(* IEC 61131-3 sources: Lasal-MCP/examples/SampleSource/4_PumpControlSchemeSolution/Stations/MachineControl/MachineControl/Class/_EventAddfromPLC, 1 file *)

(* ---- _EventAddfromPLC.st ---- *)
#ifndef EVENT_VALUECHANGE
  #define   Event_ValueChange               16#102      // Event für: Variable vom Typ Numeric
#endif

#ifndef EVENT_EVENTENTRY
  #define   Event_EventEntry                16#270
#endif

(*!
<Class
	Name               = "_EventAddfromPLC"
	Revision           = "1.4"
	RealtimeTask       = "false"
	CyclicTask         = "true"
	BackgroundTask     = "true"
	Sigmatek           = "true"
	OSInterface        = "false"
	HighPriority       = "false"
	Automatic          = "false"
	UpdateMode         = "Prescan"
	SharedCommandTable = "true"
	Objectsize         = "(470,120)"
	Comment            = "class for adding an event from plc and sending it to HMI via DataManager">
	<Channels>
		<Server Name="ClassSvr">
			<NewInst>
				<Function Name="NewInst_AddSystemOnOff">
					<InputParameter>
						<Parameter Name="dDate"/>
						<Parameter Name="dTime"/>
						<Parameter Name="bSwitchOnOff"/>
					</InputParameter>
					<OutputParameter>
						<Parameter Name="ret_code"/>
					</OutputParameter>
				</Function>
				<Function Name="NewInst_AddEventEntry">
					<InputParameter>
						<Parameter Name="config"/>
						<Parameter Name="uiCategory"/>
						<Parameter Name="uiIndex"/>
						<Parameter Name="pText"/>
						<Parameter Name="uiSize"/>
						<Parameter Name="bUnicode"/>
					</InputParameter>
					<OutputParameter>
						<Parameter Name="ret_code"/>
					</OutputParameter>
				</Function>
				<Function Name="NewInst_AddDateChange">
					<InputParameter>
						<Parameter Name="udVarNo"/>
						<Parameter Name="dOldDate"/>
						<Parameter Name="dNewDate"/>
					</InputParameter>
					<OutputParameter>
						<Parameter Name="ret_code"/>
					</OutputParameter>
				</Function>
				<Function Name="NewInst_AddTimeChange">
					<InputParameter>
						<Parameter Name="udVarNo"/>
						<Parameter Name="dOldTime"/>
						<Parameter Name="dNewTime"/>
					</InputParameter>
					<OutputParameter>
						<Parameter Name="ret_code"/>
					</OutputParameter>
				</Function>
				<Function Name="NewInst_AddMenuChange">
					<InputParameter>
						<Parameter Name="udVarNo"/>
						<Parameter Name="udMenuIndex"/>
						<Parameter Name="dOldValue"/>
						<Parameter Name="dNewValue"/>
					</InputParameter>
					<OutputParameter>
						<Parameter Name="ret_code"/>
					</OutputParameter>
				</Function>
				<Function Name="NewInst_AddValueChange">
					<InputParameter>
						<Parameter Name="udLasalID"/>
						<Parameter Name="dOldValue"/>
						<Parameter Name="dNewValue"/>
					</InputParameter>
					<OutputParameter>
						<Parameter Name="ret_code"/>
					</OutputParameter>
				</Function>
				<Function Name="NewInst_AddOPChange">
					<InputParameter>
						<Parameter Name="eOPMode"/>
					</InputParameter>
					<OutputParameter>
						<Parameter Name="ret_code"/>
					</OutputParameter>
				</Function>
				<Function Name="NewInst_AddUserLoginLogout">
					<InputParameter>
						<Parameter Name="pUserName"/>
						<Parameter Name="dActLevel"/>
						<Parameter Name="bIsLogin"/>
					</InputParameter>
					<OutputParameter>
						<Parameter Name="ret_code"/>
					</OutputParameter>
				</Function>
			</NewInst>
		</Server>
	</Channels>
	<Dependencies>
		<Files>
			<File Path=".\Class\_EventAddfromPLC\_EventAddfromPLC_de.pdf"/>
			<File Path=".\Class\_EventAddfromPLC\_EventAddfromPLC_en.pdf"/>
		</Files>
	</Dependencies>
	<RevDoku>
		<Owner Company="Sigmatek"/>
		<Dokumentation Revision="1.4" Date="2016-10-21" Author="KaiAnd" Company="Sigmatek" Description="implemented NewInst_AddXY (Cmd 00 to Cmd 07) for adding events from external via command channel"/>
		<Dokumentation Revision="1.3" Date="2016-10-10" Author="HubChr" Company="Sigmatek" Description="Added documentation pdfs."/>
		<Dokumentation Revision="1.2" Date="2016-09-21" Author="HubChr" Company="Sigmatek" Description="Events from PLC can now also open MessageBoxes"/>
		<Dokumentation Revision="1.1" Date="2016-09-15" Author="HubChr" Company="Sigmatek" Description="Translated comments for library compatibility"/>
		<Dokumentation Revision="1.0" Date="2015-09-22" Company="Sigmatek" Description="Creation."/>
	</RevDoku>
	<Network Name="_EventAddfromPLC">
		<!-- List of Components in this network -->
		<Components>
			<Object
				Name       = "_base"
				Class      = "TCPComSend"
				Position   = "(218,120)"
				Visualized = "false">
				<Channels>
					<Server Name="ClassSvr"/>
					<Server Name="ID_Destination"/>
					<Server Name="ID_Source"/>
					<Server Name="sSendCnt"/>
					<Server Name="sSendErr"/>
					<Client Name="cPrio"/>
					<Client Name="cSendErr"/>
					<Client Name="cSendOk"/>
					<Client Name="toDataManager"/>
				</Channels>
			</Object>
		</Components>
		<Comments>
		</Comments>
		<!-- List of Connections in this network -->
		<Connections>
			<Connection Source="this.ClassSvr" Destination="_base.ClassSvr" Vertices="(1006,210),(834,210),"/>
			<Connection Source="this.ID_Destination" Destination="_base.ID_Destination" Vertices="(1006,270),(834,270),"/>
			<Connection Source="this.ID_Source" Destination="_base.ID_Source" Vertices="(1006,330),(834,330),"/>
			<Connection Source="this.sSendCnt" Destination="_base.sSendCnt" Vertices="(1006,390),(834,390),"/>
			<Connection Source="this.sSendErr" Destination="_base.sSendErr" Vertices="(1006,450),(834,450),"/>
			<Connection Source="_base.toDataManager" Destination="this.toDataManager" Vertices="(218,210),(38,210),"/>
			<Connection Source="_base.cPrio" Destination="this.cPrio" Vertices="(218,270),(38,270),"/>
		</Connections>
		<!-- Headerfiles -->
		<Options>
		</Options>
	</Network>
</Class>
*)
#pragma using TCPComSend

_EventAddfromPLC : CLASS
: TCPComSend
	TYPE
#pragma pack(push, 1)
	  _PLCEventdata : STRUCT
	    EventType : UINT;
	    no_para : UINT;
	    Para1 : DINT;
	    Para2 : DINT;
	    Para3 : DINT;
	    Para4 : DINT;
	    Para5 : DINT;
	    Para6 : DINT;
	    Para7 : DINT;
	    Para8 : DINT;
	    StringSize : UINT;
	    aString : ARRAY [0..24] OF DINT;
	  END_STRUCT;
#pragma pack(pop)
	  CmdClassSvr :  //! <Type Public="true" Name="CmdClassSvr"/>
	  (
	    NewInst_AddSystemOnOff:=0,
	    NewInst_AddEventEntry,
	    NewInst_AddDateChange,
	    NewInst_AddTimeChange,
	    NewInst_AddMenuChange,
	    NewInst_AddValueChange,
	    NewInst_AddOPChange,
	    NewInst_AddUserLoginLogout
	  )$UINT;
	END_TYPE
  //Servers:
  //Clients:
  //Variables:
  //Functions:
				//! <Function Comment="Initialization of the eventdata." Name="InitPLCEventdata"/>
	FUNCTION InitPLCEventdata
		VAR_INPUT
			pPLCEvent 	: ^_PLCEventdata;			//! <Variable Comment="Pointer to the event data." Name="InitPLCEventdata.pPLCEvent"/>
		END_VAR;
				//! <Function Comment="Sends an event for a value change to the remote station." Name="AddValueChange"/>
	FUNCTION GLOBAL AddValueChange
		VAR_INPUT
			udLasalID 	: UDINT;			//! <Variable Comment="Lasal-ID" Name="AddValueChange.udLasalID"/>
			dOldValue 	: DINT;			//! <Variable Comment="Old value" Name="AddValueChange.dOldValue"/>
			dNewValue 	: DINT;			//! <Variable Comment="New value" Name="AddValueChange.dNewValue"/>
		END_VAR;
				//! <Function Comment="Method for sending the data of a event to the remote station." Name="AddEventEntry"/>
	FUNCTION GLOBAL AddEventEntry
		VAR_INPUT
			config 	: BDINT;			//! <Variable Comment="Category for the event:&#13;&#10;0 .. System category 1&#13;&#10;1 .. System category 2&#13;&#10;2 .. System category 3&#13;&#10;3 .. System category 4&#13;&#10;4 .. Change of the OP mode&#13;&#10;else .. System category 1" Name="AddEventEntry.config"/>
			uiCategory 	: UINT;			//! <Variable Comment="Category for the event:&#13;&#10;0 .. System category 1&#13;&#10;1 .. System category 2&#13;&#10;2 .. System category 3&#13;&#10;3 .. System category 4&#13;&#10;4 .. Change of the OP mode&#13;&#10;else .. System category 1" Name="AddEventEntry.uiCategory"/>
			uiIndex 	: UINT;			//! <Variable Comment="Index in the textscheme (if used).&#13;&#10;Note: If event is for example a menue-change -&gt; menue-index." Name="AddEventEntry.uiIndex"/>
			pText 	: ^void;			//! <Variable Comment="Individual text" Name="AddEventEntry.pText"/>
			uiSize 	: UINT;			//! <Variable Comment="Size of the text" Name="AddEventEntry.uiSize"/>
			bUnicode 	: BOOL;			//! <Variable Comment="Character size of the string:&#13;&#10;FALSE .. ASCII&#13;&#10;TRUE .. UNI-Code" Name="AddEventEntry.bUnicode"/>
		END_VAR;

	FUNCTION ClassSvr::NewInst_AddSystemOnOff
		VAR_INPUT
			dDate 	: DINT;
			dTime 	: DINT;
			bSwitchOnOff 	: DINT;
		END_VAR
		VAR_OUTPUT
			ret_code 	: IprStates;
		END_VAR;

	FUNCTION ClassSvr::NewInst_AddEventEntry
		VAR_INPUT
			config 	: DINT;
			uiCategory 	: DINT;
			uiIndex 	: DINT;
			pText 	: DINT;
			uiSize 	: DINT;
			bUnicode 	: DINT;
		END_VAR
		VAR_OUTPUT
			ret_code 	: IprStates;
		END_VAR;

	FUNCTION ClassSvr::NewInst_AddDateChange
		VAR_INPUT
			udVarNo 	: DINT;
			dOldDate 	: DINT;
			dNewDate 	: DINT;
		END_VAR
		VAR_OUTPUT
			ret_code 	: IprStates;
		END_VAR;

	FUNCTION ClassSvr::NewInst_AddTimeChange
		VAR_INPUT
			udVarNo 	: DINT;
			dOldTime 	: DINT;
			dNewTime 	: DINT;
		END_VAR
		VAR_OUTPUT
			ret_code 	: IprStates;
		END_VAR;

	FUNCTION ClassSvr::NewInst_AddMenuChange
		VAR_INPUT
			udVarNo 	: DINT;
			udMenuIndex 	: DINT;
			dOldValue 	: DINT;
			dNewValue 	: DINT;
		END_VAR
		VAR_OUTPUT
			ret_code 	: IprStates;
		END_VAR;

	FUNCTION ClassSvr::NewInst_AddValueChange
		VAR_INPUT
			udLasalID 	: DINT;
			dOldValue 	: DINT;
			dNewValue 	: DINT;
		END_VAR
		VAR_OUTPUT
			ret_code 	: IprStates;
		END_VAR;

	FUNCTION ClassSvr::NewInst_AddOPChange
		VAR_INPUT
			eOPMode 	: DINT;
		END_VAR
		VAR_OUTPUT
			ret_code 	: IprStates;
		END_VAR;

	FUNCTION ClassSvr::NewInst_AddUserLoginLogout
		VAR_INPUT
			pUserName 	: DINT;
			dActLevel 	: DINT;
			bIsLogin 	: DINT;
		END_VAR
		VAR_OUTPUT
			ret_code 	: IprStates;
		END_VAR;
				//! <Function Name="ClassSvr.NewInst" Hidden="true"/>
	FUNCTION VIRTUAL GLOBAL ClassSvr::NewInst
		VAR_INPUT
			pPara 	: ^CmdStruct;
			pResult 	: ^results;
		END_VAR
		VAR_OUTPUT
			ret_code 	: iprStates;
		END_VAR;
  //Tables:
	FUNCTION @STD
		VAR_OUTPUT
			ret_code	: CONFSTATES;
		END_VAR;
	FUNCTION GLOBAL TAB @CT_;
END_CLASS;

FUNCTION VIRTUAL GLOBAL _EventAddfromPLC::ClassSvr::NewInst
	VAR_INPUT
		pPara 	: ^CmdStruct;
		pResult 	: ^Results;
	END_VAR
	VAR_OUTPUT
		ret_code 	: IprStates;
	END_VAR
	CASE pPara^.uiCmd$CmdClassSvr OF
		NewInst_AddSystemOnOff:
			ret_code := NewInst_AddSystemOnOff(pPara^.aPara[0],pPara^.aPara[1],pPara^.aPara[2]);
			pResult^.uiLng := 0 + sizeof(pResult^.uiLng);
		NewInst_AddEventEntry:
			ret_code := NewInst_AddEventEntry(pPara^.aPara[0],pPara^.aPara[1],pPara^.aPara[2],pPara^.aPara[3],pPara^.aPara[4],pPara^.aPara[5]);
			pResult^.uiLng := 0 + sizeof(pResult^.uiLng);
		NewInst_AddDateChange:
			ret_code := NewInst_AddDateChange(pPara^.aPara[0],pPara^.aPara[1],pPara^.aPara[2]);
			pResult^.uiLng := 0 + sizeof(pResult^.uiLng);
		NewInst_AddTimeChange:
			ret_code := NewInst_AddTimeChange(pPara^.aPara[0],pPara^.aPara[1],pPara^.aPara[2]);
			pResult^.uiLng := 0 + sizeof(pResult^.uiLng);
		NewInst_AddMenuChange:
			ret_code := NewInst_AddMenuChange(pPara^.aPara[0],pPara^.aPara[1],pPara^.aPara[2],pPara^.aPara[3]);
			pResult^.uiLng := 0 + sizeof(pResult^.uiLng);
		NewInst_AddValueChange:
			ret_code := NewInst_AddValueChange(pPara^.aPara[0],pPara^.aPara[1],pPara^.aPara[2]);
			pResult^.uiLng := 0 + sizeof(pResult^.uiLng);
		NewInst_AddOPChange:
			ret_code := NewInst_AddOPChange(pPara^.aPara[0]);
			pResult^.uiLng := 0 + sizeof(pResult^.uiLng);
		NewInst_AddUserLoginLogout:
			ret_code := NewInst_AddUserLoginLogout(pPara^.aPara[0],pPara^.aPara[1],pPara^.aPara[2]);
			pResult^.uiLng := 0 + sizeof(pResult^.uiLng);
	ELSE

	ret_code := READY;
	END_CASE;

END_FUNCTION

FUNCTION _EventAddfromPLC::InitPLCEventdata
	VAR_INPUT
		pPLCEvent 	: ^_PLCEventdata;
	END_VAR

  pPLCEvent^.EventType  := 0;
  pPLCEvent^.no_para    := 0;
  pPLCEvent^.Para1      := 0;
  pPLCEvent^.Para2      := 0;
  pPLCEvent^.Para3      := 0;
  pPLCEvent^.Para4      := 0;
  pPLCEvent^.Para5      := 0;
  pPLCEvent^.Para6      := 0;
  pPLCEvent^.Para7      := 0;
  pPLCEvent^.Para8      := 0;
  pPLCEvent^.StringSize := 0;
  _memset(dest := #pPLCEvent^.aString[0], usByte:=0, cntr:=sizeof(pPLCEvent^.aString));

END_FUNCTION

FUNCTION GLOBAL _EventAddfromPLC::AddValueChange
	VAR_INPUT
		udLasalID : UDINT;
		dOldValue : DINT;
		dNewValue : DINT;
	END_VAR
  VAR
  	tmpEvent : _PLCEventdata;
  END_VAR

  InitPLCEventdata(pPLCEvent:=#tmpEvent);

  // add event for change of value
  tmpEvent.EventType := EVENT_VALUECHANGE;

  // store information
  tmpEvent.no_para := 3;
  tmpEvent.para1   := udLasalID$DINT;
  tmpEvent.para2   := dOldValue;
  tmpEvent.para3   := dNewValue;

  SendData(pData:=#tmpEvent$^void, length:=sizeof(tmpEvent), timeout:=1000, OptCMD:=0);

END_FUNCTION

FUNCTION GLOBAL _EventAddfromPLC::AddEventEntry
	VAR_INPUT
		config 	   : BDINT;
		uiCategory : UINT;
		uiIndex 	 : UINT;
		pText 	   : ^void;
		uiSize 	   : UINT;
		bUnicode 	 : BOOL;
	END_VAR
  VAR
  	tmpEvent : _PLCEventdata;
  END_VAR

  InitPLCEventdata(pPLCEvent:=#tmpEvent);

  tmpEvent.EventType := EVENT_EVENTENTRY;

  // store information
  tmpEvent.no_para := 3;
  tmpEvent.para1   := to_dint(uiCategory);
  tmpEvent.para2   := to_dint(uiIndex);
  tmpEvent.para3   := bUnicode;
  tmpEvent.para4   := config$DINT;

  if ( (pText <> NIL) & (uiSize < (sizeof(tmpEvent.aString) -1)) ) then

    tmpEvent.StringSize := uiSize;
    _memcpy(ptr1:=#tmpEvent.aString[0], ptr2:=pText, cntr:=uiSize);

  end_if;

  SendData(pData:=#tmpEvent$^void, length:=sizeof(tmpEvent), timeout:=1000, OptCMD:=0);

END_FUNCTION

//***********************************************************************************************************
//  NewInst Commands for external actions via command channel
//***********************************************************************************************************

//-------------------------------------------------------------------------------------------------
//  Cmd 00: AddSystemOnOff
//-------------------------------------------------------------------------------------------------
#pragma warning(disable:73);
FUNCTION _EventAddfromPLC::NewInst_AddSystemOnOff
	VAR_INPUT
		dDate 	: DINT;
		dTime 	: DINT;
		bSwitchOnOff 	: DINT;
	END_VAR
	VAR_OUTPUT
		ret_code 	: IprStates;
	END_VAR

	ret_code := READY;

// NOT IMPLEMENTED IN PLC - reserverd for future

//  AddSystemOnOff( dDate        := dDate,
//                  dTime        := dTime,
//                  bSwitchOnOff := TO_BOOL(bSwitchOnOff) );

END_FUNCTION
#pragma warning(default:73);

//-------------------------------------------------------------------------------------------------
//  Cmd 01: AddEventEntry
//-------------------------------------------------------------------------------------------------
FUNCTION _EventAddfromPLC::NewInst_AddEventEntry
	VAR_INPUT
		config 	: DINT;
		uiCategory 	: DINT;
		uiIndex 	: DINT;
		pText 	: DINT;
		uiSize 	: DINT;
		bUnicode 	: DINT;
	END_VAR
	VAR_OUTPUT
		ret_code 	: IprStates;
	END_VAR

	ret_code := READY;

  AddEventEntry(config     := config$BDINT,
                uiCategory := TO_UINT(uiCategory),
                uiIndex    := TO_UINT(uiIndex),
                pText      := pText$^void,
                uiSize     := TO_UINT(uiSize),
                bUnicode   := TO_BOOL(bUnicode) );

END_FUNCTION

//-------------------------------------------------------------------------------------------------
//  Cmd 02: AddDateChange
//-------------------------------------------------------------------------------------------------
#pragma warning(disable:73);
FUNCTION _EventAddfromPLC::NewInst_AddDateChange
	VAR_INPUT
		udVarNo 	: DINT;
		dOldDate 	: DINT;
		dNewDate 	: DINT;
	END_VAR
	VAR_OUTPUT
		ret_code 	: IprStates;
	END_VAR

	ret_code := READY;

// NOT IMPLEMENTED IN PLC - reserverd for future

//  AddDateChange(udVarNo  := udVarNo$UDINT,
//                dOldDate := dOldDate,
//                dNewDate := dNewDate );

END_FUNCTION
#pragma warning(default:73);

//-------------------------------------------------------------------------------------------------
//  Cmd 03: AddTimeChange
//-------------------------------------------------------------------------------------------------
#pragma warning(disable:73);
FUNCTION _EventAddfromPLC::NewInst_AddTimeChange
	VAR_INPUT
		udVarNo 	: DINT;
		dOldTime 	: DINT;
		dNewTime 	: DINT;
	END_VAR
	VAR_OUTPUT
		ret_code 	: IprStates;
	END_VAR

	ret_code := READY;

// NOT IMPLEMENTED IN PLC - reserverd for future

//  AddTimeChange(udVarNo  := udVarNo$UDINT,
//                dOldTime := dOldTime,
//                dNewTime := dNewTime );

END_FUNCTION
#pragma warning(default:73);

//-------------------------------------------------------------------------------------------------
//  Cmd 04: AddMenuChange
//-------------------------------------------------------------------------------------------------
#pragma warning(disable:73);
FUNCTION _EventAddfromPLC::NewInst_AddMenuChange
	VAR_INPUT
		udVarNo 	: DINT;
		udMenuIndex 	: DINT;
		dOldValue 	: DINT;
		dNewValue 	: DINT;
	END_VAR
	VAR_OUTPUT
		ret_code 	: IprStates;
	END_VAR

	ret_code := READY;

// NOT IMPLEMENTED IN PLC - reserverd for future

//  AddMenuChange(udVarNo     := udVarNo$UDINT,
//                udMenuIndex := udMenuIndex$UDINT,
//                dOldValue   := dOldValue,
//                dNewValue   := dNewValue );

END_FUNCTION
#pragma warning(default:73);

//-------------------------------------------------------------------------------------------------
//  Cmd 05: AddValueChange
//-------------------------------------------------------------------------------------------------
FUNCTION _EventAddfromPLC::NewInst_AddValueChange
	VAR_INPUT
		udLasalID : DINT;
		dOldValue : DINT;
		dNewValue : DINT;
	END_VAR
	VAR_OUTPUT
		ret_code 	: IprStates;
	END_VAR

	ret_code := READY;

  AddValueChange( udLasalID := udLasalID$UDINT,
                  dOldValue := dOldValue,
                  dNewValue := dNewValue );

END_FUNCTION

//-------------------------------------------------------------------------------------------------
//  Cmd 06: AddOPChange
//-------------------------------------------------------------------------------------------------
#pragma warning(disable:73);
FUNCTION _EventAddfromPLC::NewInst_AddOPChange
	VAR_INPUT
		eOPMode 	: DINT;
	END_VAR
	VAR_OUTPUT
		ret_code 	: IprStates;
	END_VAR

	ret_code := READY;

// NOT IMPLEMENTED IN PLC - reserverd for future

//  AddOPChange(eOPMode := eOPMode$t_e_OPMode);

END_FUNCTION
#pragma warning(default:73);

//-------------------------------------------------------------------------------------------------
//  Cmd 07: AddUserLoginLogout
//-------------------------------------------------------------------------------------------------
#pragma warning(disable:73);
FUNCTION _EventAddfromPLC::NewInst_AddUserLoginLogout
	VAR_INPUT
		pUserName 	: DINT;
		dActLevel 	: DINT;
		bIsLogin 	: DINT;
	END_VAR
	VAR_OUTPUT
		ret_code 	: IprStates;
	END_VAR

	ret_code := READY;

// NOT IMPLEMENTED IN PLC - reserverd for future

//  AddUserLoginLogout( pUserName := pUserName$^CHAR,
//                      dActLevel := dActLevel,
//                      bIsLogin  := TO_BOOL(bIsLogin) );

END_FUNCTION
#pragma warning(default:73);

//***********************************************************************************************************
